(*
SPDX-FileCopyrightText: © 2026 Oleksandr Tiutyk <trofimich@gmail.com>
SPDX-License-Identifier: MIT
License: https://opensource.org/license/mit
*)

(*!
<summary>
Beckhoff EL5001: 1-channel SSI absolute encoder interface terminal.
</summary>
<description>
Process image mapping structure for the EL5001 synchronous serial interface (SSI) absolute encoder terminal.
Requires firmware 11 or later and the two-byte status PDO 0x1A01. The one-byte variant is unsupported.
When used for I/O, link located fields or their containing buffers to the matching selected PDOs.
The record is not a packed wire buffer; compiler padding is not part of the device specification.
Unlinked/default values do not prove valid I/O. The caller evaluates bus/channel validity before use.
Use one owner task per instance and externally synchronize other access; multi-field snapshots are not atomic.
Copies store data without creating hardware links. Keep borrowed field references valid while consumers are bound.
This passive record performs no validation, synchronization, configuration or protocol advancement.
</description>
*)
TYPE EL5001 :
STRUCT
	Ch1 : SSI_ENCODER_CHANNEL;
END_STRUCT
END_TYPE

(* stored: Version 1.1.0.1, ProductVersion 3.1.4026.20
   DUT EL5001: Id {b0179e9e-88ae-4c6e-9fed-4547d54ae337} *)
